# EPICS StreamDevice protocol: EPICS/Db/tic.proto
# tic.proto - Edwards TIC controller over RS-232 (databases: tic.db, task T29; tic_control.db, T32)
#
# The protocols down to "ident_sw" are queries only, and they are all that tic.db uses: tic.db
# alone sends no command ("!C") and no setup ("!S"). The protocols at the end ("command", task T32)
# send a command; only tic_control.db uses them, for the requests of the station's two pumps and
# of one gauge. No protocol here sends a setup ("!S").
#
# Source: Edwards "Turbo Instrument Controller (TIC) Serial Communications", D397-30-880 Issue H
# (2012), which covers all seven TIC variants (Instrument Controller 3 and 6 gauges, Turbo
# Controller, Turbo & Instrument Controller):
#   1.2    query "?V<obj>" / "?S<obj>", every message ends with CR, the TIC answers only when asked
#   1.6    replies "=V<obj> <data>" / "=S<obj> <data>" or the response code "*V<obj> <r>" /
#          "*S<obj> <r>" (Table 3); fields of the data separated by ";" (1.5)
#   1.4    basic messages answered in less than 100 ms; suggested master timeout 500 ms
#   Table 1, 1.6.2.2, 1.6.2.3: the objects below
# Every reply names its object, so a late reply to another query cannot be taken for this one.
#
# ReplyTimeout 150 ms, not the 500 ms the manual suggests: with 500 ms one silent cycle would
# need 6.6 s of line time every 2 s. Seen on the lab's controller on 2026-11-25 (the probe, a
# Prolific adapter): replies after 23 to 50 ms, the identity after 61 and 86 ms. 150 ms leaves
# 64 ms on the slowest, and 13 queries of a silent controller take 1.95 s of the 2 s (120 ms,
# from the manual's "less than 100 ms", was the value before the measurement). None of these
# queries is routed to a DX/nEXT pump (objects 800+, 200 ms). Line budget: docs/emulation/TIC.md.
#
# The records of the value queries are calcout records: StreamDevice writes the fields of the
# reply into the record's own fields A, B, C ... (%(A) etc., no processing), the error code of an
# error reply into F. The record's CALC sets these fields to "nothing" (NAN, -1) before every
# request, so no field keeps a value of an earlier reply. An error reply leaves the record in
# INVALID/CALC (the @mismatch handler of StreamDevice), a missing one in INVALID/TIMEOUT.

Terminator = CR;
ReplyTimeout = 150;
ReadTimeout = 50;

# Gauge 1, 2, 3 (objects 913, 914, 915; Table 1): "?V913" -> "=V913 value;units type;state;
# alert ID;priority". Value: pressure in pascal when units type is 59 (1.7.4: "PRESSURE 59 -
# float (Pascals only)"), volts when 66. State: 1.7.7. Alert: 1.7.3. Priority: 1.7.2.
gauge {
    out "?V\$1";
    in "=V\$1 %(A)g;%(B)d;%(C)d;%(D)d;%(E)d";
    @mismatch { in "*V\$1 %(F)d"; }
}

# Turbo pump (904, 1.6.2.3) and backing pump (910, Table 1): "state;alert ID;priority".
# Turbo states: 1.7.8 "Full pump states" 0-7. Backing: "State 0 - 4" (Table 1), the states of 1.7.6.
pump {
    out "?V\$1";
    in "=V\$1 %(A)d;%(B)d;%(C)d";
    @mismatch { in "*V\$1 %(F)d"; }
}

# Turbo speed (905, Table 1): "value;alert ID;priority", value 0.0 - 110.0 %.
speed {
    out "?V\$1";
    in "=V\$1 %(A)g;%(B)d;%(C)d";
    @mismatch { in "*V\$1 %(F)d"; }
}

# Pump type (904, 910): query setup with config type 3, "?S904 3" -> "=S904 3;p" (1.6.2.3,
# Table 1), p from 1.7.11 (0 = No Pump).
pump_type {
    out "?S\$1 3";
    in "=S\$1 3;%(A)d";
    @mismatch { in "*S\$1 %(F)d"; }
}

# System status (902 ?V, Table 1): one state value per item, then alert ID and priority. The
# number of fields depends on the variant: TC 7, IC 8, TIC 10, IC6 14 (aai record, NORD).
system {
    Separator = ";";
    out "?V902";
    in "=V902 %d";
}

# Identity (902 ?S, 1.6.2.2): "TIC;Dxxxxxxxx;serial number;PIC s/w ver", max 80 characters.
# The lab's controller answers '=S902 TIC100;D39700640T;160070509<00>;5.0' (seen 2026-11-25):
# a NUL byte after the serial number. The text conversion ends at the NUL, and without
# ExtraInput = Ignore the rest ("<00>;5.0") is surplus input and the record INVALID (seen with
# the simulator sending this form). So the identity is type, software and serial number; the
# PIC software version behind the NUL is not read.
ident {
    ExtraInput = Ignore;
    out "?S902";
    in "=S902 %80[^\r]";
}

# The first two fields of every identity reply that ident requested (SCAN I/O Intr: they send
# nothing). They keep their last value while the controller is silent; ident:get then is INVALID.
ident_model {
    ExtraInput = Ignore;
    in "=S902 %39[^;]";
}
ident_sw {
    ExtraInput = Ignore;
    in "=S902 %*[^;];%39[^;]";
}

# ------------------------------------------------------------------ task T32 (tic_control.db)

# A command: "!C<obj> <d>", answered "*C<obj> <r>" (D397-30-880 Table 1: 904 turbo pump and 910
# backing pump "Turn pump on/off", On = 1, Off = 0; 913-915 gauges "On/off", 1.7.5 Gauge On = 1,
# Gauge Off = 0; the response codes of Table 3, 0 "no error"). Used by the request records (bo)
# of tic_control.db: the record's value is sent (%d, the RVAL of a bo without MASK: 0 or 1).
# Seen on the lab's controller (2026-11-25, sent by hand): "!C910 1", "!C910 0", "!C904 1",
# "!C904 0", each answered "*C9xx 0" after 19 ms. The gauge's "!C914 1" / "!C914 0" were not
# tried: from the manual only.
# The acknowledgement "*C<obj> 0" ends the request without alarm. Another code: the @mismatch
# handler stores it in the bo's own field IVOV (not used otherwise: the records have IVOA "Don't
# drive outputs") and the record ends INVALID/CALC; tic_control.db shows the code's word. No
# reply: INVALID/TIMEOUT. Every reply names its object, so a late reply to a query is not taken
# for the acknowledgement.
command {
    out "!C\$1 %d";
    in "*C\$1 0";
    @mismatch { in "*C\$1 %(IVOV)d"; }
}

# The slave setup of a gauge, read only: "?S<obj> 4" (Table 1, objects 913-915, config type 4:
# "Read slave setup - master; units type; on setpoint; off setpoint, enable"; master an object
# ID, gauge 1/2/3 or the turbo speed; set points in pascal for units 59). The form of the reply is
# that seen on the lab's controller for the turbopump's object 904 (2026-11-25):
# "=S904 4;0;59;0.0000e+00;0.0000e+00;0", config type first. The gauges' replies were not seen;
# the manual's own example (1.6.2.3) has no config type ("=S904 913;59;5.1e-2;4.9e-1;1"): such a
# reply, or any other form, leaves the record INVALID (CALC, as a mismatch) and slave_raw keeps
# its text. Fields into the calcout's A (master), B (units type), C (on), D (off), E (enable),
# an error code into F.
slave {
    out "?S\$1 4";
    in "=S\$1 4;%(A)d;%(B)d;%(C)g;%(D)g;%(E)d";
    @mismatch { in "*S\$1 %(F)d"; }
}

# The text of every "=S<obj> ..." reply that slave requested (SCAN I/O Intr: it sends nothing),
# whatever its form, for the first contact with a controller whose replies are not known.
slave_raw {
    ExtraInput = Ignore;
    in "=S\$1 %39[^\r]";
}
